PROGRAM ValueFactory
VAR CONSTANT
	nSpanIdBytes: USINT := 8;
	nTraceIdBytes: USINT := 16;
END_VAR

METHOD cloneAnyValue : BOOL
VAR_IN_OUT
	pDest: POINTER TO FB_AnyValue;
END_VAR
VAR_INPUT
	pSrc: POINTER TO FB_AnyValue;
END_VAR
VAR_OUTPUT
	failureReason: E_ValueFactoryFailureReason;
END_VAR
VAR
	_type: E_ValueType;
END_VAR
cloneAnyValue := FALSE;
failureReason := E_ValueFactoryFailureReason.NA;

IF pDest <> 0 THEN
	failureReason := E_ValueFactoryFailureReason.DESTINATION_ALREADY_ASSIGNED;
	RETURN;
END_IF

IF pSrc = 0 THEN
	failureReason := E_ValueFactoryFailureReason.SOURCE_POINTER_NULL;
	RETURN;
END_IF

_type := pSrc^.eType;
CASE _type OF
	E_ValueType.E_String:
		cloneAnyValue := ValueFactory.cloneString(pDest:=pDest, pSrc:=pSrc, failureReason=>failureReason);
	E_ValueType.E_Number:
		cloneAnyValue := ValueFactory.cloneNumber(pDest:=pDest, pSrc:=pSrc, failureReason=>failureReason);
	E_ValueType.E_KeyValue:
		cloneAnyValue := ValueFactory.cloneKeyValue(pDest:=pDest, pSrc:=pSrc, failureReason=>failureReason);
	ELSE
		failureReason := E_ValueFactoryFailureReason.UNSUPPORTED_VALUE_TYPE;
END_CASE
END_METHOD

METHOD cloneKeyValue : BOOL
VAR_IN_OUT
	pDest: POINTER TO FB_KeyValue;
END_VAR
VAR_INPUT
	pSrc: POINTER TO FB_KeyValue;
END_VAR
VAR_OUTPUT
	failureReason: E_ValueFactoryFailureReason;
END_VAR
cloneKeyValue := FALSE;
failureReason := E_ValueFactoryFailureReason.NA;

IF pDest <> 0 THEN
	failureReason := E_ValueFactoryFailureReason.DESTINATION_ALREADY_ASSIGNED;
	RETURN;
END_IF

IF pSrc = 0 THEN
	failureReason := E_ValueFactoryFailureReason.SOURCE_POINTER_NULL;
	RETURN;
END_IF

cloneKeyValue := ValueFactory.createKeyValue(
	pDest:=pDest,
	pKey:=pSrc^.pKey,
	pVal:=pSrc^.pVal,
	failureReason=>failureReason
);
END_METHOD

METHOD cloneNumber : BOOL
VAR_IN_OUT
	pDest: POINTER TO FB_Number;
END_VAR
VAR_INPUT
	pSrc: POINTER TO FB_Number;
END_VAR
VAR_OUTPUT
	failureReason: E_ValueFactoryFailureReason;
END_VAR
VAR
	_value: AnyType;
	_pNew: POINTER TO FB_Number;
END_VAR
cloneNumber := FALSE;
failureReason := E_ValueFactoryFailureReason.NA;

IF pDest <> 0 THEN
	failureReason := E_ValueFactoryFailureReason.DESTINATION_ALREADY_ASSIGNED;
	RETURN;
END_IF

IF pSrc = 0 THEN
	failureReason := E_ValueFactoryFailureReason.SOURCE_POINTER_NULL;
	RETURN;
END_IF

IF pSrc^.value.pValue = 0 THEN
	failureReason := E_ValueFactoryFailureReason.NUMBER_VALUE_POINTER_NULL;
	RETURN;
END_IF

IF pSrc^.value.diSize <= 0 THEN
	failureReason := E_ValueFactoryFailureReason.NUMBER_VALUE_SIZE_INVALID;
	RETURN;
END_IF

// because it's really verbose to extract the number back out of the number we manually clone numbers
_value := pSrc^.value;
_value.pValue := __NEW(BYTE, _value.diSize);
IF _value.pValue = 0 THEN
	failureReason := E_ValueFactoryFailureReason.MEMORY_ALLOCATION_FAILURE;
	RETURN;
END_IF
MEMCPY(_value.pValue, pSrc^.value.pValue, TO_UDINT(_value.diSize));

_pNew := __NEW(FB_Number(
	value:=_value
));
IF _pNew = 0 THEN
	failureReason := E_ValueFactoryFailureReason.MEMORY_ALLOCATION_FAILURE;
	__DELETE(_value.pValue);
	_value.pValue := 0;
	RETURN;
END_IF
_value.pValue := 0;  // moved into FB_Number
pDest := _pNew;
cloneNumber := failureReason = E_ValueFactoryFailureReason.NA;
END_METHOD

METHOD cloneString : BOOL
VAR_IN_OUT
	pDest: POINTER TO FB_String;
END_VAR
VAR_INPUT
	pSrc: POINTER TO FB_String;
END_VAR
VAR_OUTPUT
	failureReason: E_ValueFactoryFailureReason;
END_VAR
cloneString := FALSE;
failureReason := E_ValueFactoryFailureReason.NA;

IF pDest <> 0 THEN
	failureReason := E_ValueFactoryFailureReason.DESTINATION_ALREADY_ASSIGNED;
	RETURN;
END_IF

IF pSrc = 0 THEN
	failureReason := E_ValueFactoryFailureReason.SOURCE_POINTER_NULL;
	RETURN;
END_IF

IF pSrc^.pString = 0 THEN
	failureReason := E_ValueFactoryFailureReason.STRING_POINTER_NULL;
	RETURN;
END_IF

cloneString := ValueFactory.createString(pDest:=pDest, pString:=pSrc^.pString, failureReason=>failureReason);
END_METHOD

METHOD createKeyValue : BOOL
VAR_IN_OUT
	pDest: POINTER TO FB_KeyValue;
END_VAR
VAR_INPUT
	pKey: POINTER TO STRING;
	pVal: POINTER TO FB_AnyValue;
END_VAR
VAR_OUTPUT
	failureReason: E_ValueFactoryFailureReason;
END_VAR
VAR
	_pNew: POINTER TO FB_KeyValue;
	_pKey: POINTER TO STRING;
	_pVal: POINTER TO FB_AnyValue;
	_len: UDINT;
END_VAR
createKeyValue := FALSE;
failureReason := E_ValueFactoryFailureReason.NA;

IF pKey = 0 THEN
	failureReason := E_ValueFactoryFailureReason.KEY_POINTER_NULL;
	RETURN;
END_IF

IF pVal = 0 THEN
	failureReason := E_ValueFactoryFailureReason.VALUE_POINTER_NULL;
	RETURN;
END_IF

IF pDest <> 0 THEN
	failureReason := E_ValueFactoryFailureReason.DESTINATION_ALREADY_ASSIGNED;
	RETURN;
END_IF

// clone all owned data before allocating the value itself
_len := LEN2(pKey) + 1;
_pKey := __NEW(BYTE, _len);
IF _pKey = 0 THEN
	failureReason := E_ValueFactoryFailureReason.MEMORY_ALLOCATION_FAILURE;
	RETURN;
END_IF
MEMCPY(_pKey, pKey, _len);

createKeyValue := ValueFactory.cloneAnyValue(pDest:=_pVal, pSrc:=pVal, failureReason=>failureReason);
IF NOT createKeyValue THEN
	__DELETE(_pKey);
	_pKey := 0;
	IF _pVal <> 0 THEN _pVal^.delete(pSelf:=_pVal); END_IF
	RETURN;
END_IF

_pNew := __NEW(FB_KeyValue(pKey:=_pKey, pVal:=_pVal));
IF _pNew = 0 THEN
	createKeyValue := FALSE;
	failureReason := E_ValueFactoryFailureReason.MEMORY_ALLOCATION_FAILURE;
	__DELETE(_pKey);
	_pKey := 0;
	_pVal^.delete(pSelf:=_pVal);
	RETURN;
END_IF
_pKey := 0;  // moved into FB_KeyValue
_pVal := 0;
pDest := _pNew;
createKeyValue := failureReason = E_ValueFactoryFailureReason.NA;
END_METHOD

METHOD createNumber : BOOL
VAR_IN_OUT
	pDest: POINTER TO FB_Number;
END_VAR
VAR_INPUT
	value: ANY_NUM;
END_VAR
VAR_OUTPUT
	failureReason: E_ValueFactoryFailureReason;
END_VAR
createNumber := FALSE;
failureReason := E_ValueFactoryFailureReason.NA;

createNumber := ValueFactory.createNumber_AnyType(
	pDest:=pDest,
	value:=value,
	failureReason=>failureReason
);
END_METHOD

(*
	This method is necessary because it makes it possible to easily create
	instance of an FB_Number from already instantiated instances of FB_Number
	i.e. cloning, when the original number is gone, but the AnyType value exists.
*)
METHOD createNumber_AnyType : BOOL
VAR_IN_OUT
	pDest: POINTER TO FB_Number;
END_VAR
VAR_INPUT
	value: AnyType;  // notice this is a struct and not the ANY_NUM keyword
END_VAR
VAR_OUTPUT
	failureReason: E_ValueFactoryFailureReason;
END_VAR
VAR
	_value: AnyType;
	_pNew: POINTER TO FB_Number;
END_VAR
createNumber_AnyType := FALSE;
failureReason := E_ValueFactoryFailureReason.NA;

IF pDest <> 0 THEN
	failureReason := E_ValueFactoryFailureReason.DESTINATION_ALREADY_ASSIGNED;
	RETURN;
END_IF

IF value.pValue = 0 THEN
	failureReason := E_ValueFactoryFailureReason.NUMBER_VALUE_POINTER_NULL;
	RETURN;
END_IF

IF value.diSize <= 0 THEN
	failureReason := E_ValueFactoryFailureReason.NUMBER_VALUE_SIZE_INVALID;
	RETURN;
END_IF

// Copy the concrete numeric value so the wrapper never retains caller-owned data.
_value.TypeClass := value.TypeClass;
_value.diSize := value.diSize;
_value.pValue := __NEW(BYTE, TO_UDINT(_value.diSize));
IF _value.pValue = 0 THEN
	failureReason := E_ValueFactoryFailureReason.MEMORY_ALLOCATION_FAILURE;
	RETURN;
END_IF
MEMCPY(_value.pValue, value.pValue, TO_UDINT(value.diSize));

_pNew := __NEW(FB_Number(value:=_value));
IF _pNew = 0 THEN
	failureReason := E_ValueFactoryFailureReason.MEMORY_ALLOCATION_FAILURE;
	__DELETE(_value.pValue);
	_value.pValue := 0;
	RETURN;
END_IF
_value.pValue := 0;  // moved into FB_Number
pDest := _pNew;
createNumber_AnyType := failureReason = E_ValueFactoryFailureReason.NA;
END_METHOD

METHOD createSpanId : BOOL
VAR_IN_OUT
	pDest: POINTER TO FB_SpanId;
END_VAR
VAR_INPUT
	pBytes: POINTER TO BYTE;
	nSize: UDINT;
END_VAR
VAR_OUTPUT
	failureReason: E_ValueFactoryFailureReason;
END_VAR
VAR
	_pNew: POINTER TO FB_SpanId;
END_VAR
createSpanId := FALSE;
failureReason := E_ValueFactoryFailureReason.NA;

IF pDest <> 0 THEN
	failureReason := E_ValueFactoryFailureReason.DESTINATION_ALREADY_ASSIGNED;
	RETURN;
END_IF

IF pBytes = 0 THEN
	failureReason := E_ValueFactoryFailureReason.SPAN_ID_BYTES_POINTER_NULL;
	RETURN;
END_IF

IF nSize < ValueFactory.nSpanIdBytes THEN
	failureReason := E_ValueFactoryFailureReason.SPAN_ID_BYTE_COUNT_TOO_SMALL;
	RETURN;
END_IF

_pNew := __NEW(FB_SpanId);
IF _pNew = 0 THEN
	failureReason := E_ValueFactoryFailureReason.MEMORY_ALLOCATION_FAILURE;
	RETURN;
END_IF

MEMCPY(ADR(_pNew^.bytes), pBytes, SIZEOF(_pNew^.bytes));
pDest := _pNew;
createSpanId := failureReason = E_ValueFactoryFailureReason.NA;
END_METHOD

METHOD createString : BOOL
VAR_IN_OUT
	pDest: POINTER TO FB_String;
END_VAR
VAR_INPUT
	pString: POINTER TO STRING;
END_VAR
VAR_OUTPUT
	failureReason: E_ValueFactoryFailureReason;
END_VAR
VAR
	_pString: POINTER TO STRING;
	_pNew: POINTER TO FB_String;
	_len: UDINT;
END_VAR
createString := FALSE;
failureReason := E_ValueFactoryFailureReason.NA;

IF pDest <> 0  THEN
	failureReason := E_ValueFactoryFailureReason.DESTINATION_ALREADY_ASSIGNED;
	RETURN;
END_IF

IF pString = 0 THEN
	failureReason := E_ValueFactoryFailureReason.STRING_POINTER_NULL;
	RETURN;
END_IF

// clone the string into a new pointer so as to not use mutable data
// an extra character is needed for the terminating character, which is a literal 0 just like "cstrings"
_len := LEN2(pString) + 1;
_pString := __NEW(BYTE, _len);
IF _pString = 0 THEN
	failureReason := E_ValueFactoryFailureReason.MEMORY_ALLOCATION_FAILURE;
	RETURN;
END_IF
MEMCPY(_pString, pString, _len);

_pNew := __NEW(FB_String(pString:=_pString));
IF _pNew = 0 THEN
	failureReason := E_ValueFactoryFailureReason.MEMORY_ALLOCATION_FAILURE;
	__DELETE(_pString);
	_pString := 0;
	RETURN;
END_IF
_pString := 0;  // moved into FB_String
pDest := _pNew;
createString := failureReason = E_ValueFactoryFailureReason.NA;
END_METHOD

METHOD createTraceId : BOOL
VAR_IN_OUT
	pDest: POINTER TO FB_TraceId;
END_VAR
VAR_INPUT
	pBytes: POINTER TO BYTE;
	nSize: UDINT;
END_VAR
VAR_OUTPUT
	failureReason: E_ValueFactoryFailureReason;
END_VAR
VAR
	_pNew: POINTER TO FB_TraceId;
END_VAR
createTraceId := FALSE;
failureReason := E_ValueFactoryFailureReason.NA;

IF pDest <> 0 THEN
	failureReason := E_ValueFactoryFailureReason.DESTINATION_ALREADY_ASSIGNED;
	RETURN;
END_IF

IF pBytes = 0 THEN
	failureReason := E_ValueFactoryFailureReason.TRACE_ID_BYTES_POINTER_NULL;
	RETURN;
END_IF

IF nSize < ValueFactory.nTraceIdBytes THEN
	failureReason := E_ValueFactoryFailureReason.TRACE_ID_BYTE_COUNT_TOO_SMALL;
	RETURN;
END_IF

_pNew := __NEW(FB_TraceId);
IF _pNew = 0 THEN
	failureReason := E_ValueFactoryFailureReason.MEMORY_ALLOCATION_FAILURE;
	RETURN;
END_IF
MEMCPY(ADR(_pNew^.bytes), pBytes, SIZEOF(_pNew^.bytes));
pDest := _pNew;
createTraceId := failureReason = E_ValueFactoryFailureReason.NA;
END_METHOD

END_PROGRAM

(* stored: Version 1.1.0.1
   POU ValueFactory: Id {d187342c-6b4d-42f2-9536-f4c1c2d2d7f1}, SpecialFunc None
   Method cloneAnyValue: Id {de7b8f5c-4e52-4385-afb8-9a7f3648c37d}
   Method cloneKeyValue: Id {a8ee2c29-a418-4ec2-8e01-8ef5052daffa}
   Method cloneNumber: Id {3de2a0de-5ee7-4e65-b88c-d438e59b12f7}
   Method cloneString: Id {11bd15c6-b673-495b-8c92-4ee038baee62}
   Method createKeyValue: Id {24aad023-b447-4a30-a636-682e068d33e5}
   Method createNumber: Id {3bcb96ce-f273-4452-a75d-ea53e63d4d25}
   Method createNumber_AnyType: Id {7e7ce9b0-0c62-4b23-bdea-24531261b359}
   Method createSpanId: Id {8c55c398-28af-4759-b54f-4b55d341d11a}
   Method createString: Id {c9d254c2-678b-419f-ac3c-e884e66c3532}
   Method createTraceId: Id {34de56b8-186c-4fd3-a48c-783b8c21d02f} *)
